Yaskawa INFORM job: LAB3-GROUPV2'2.JBI

/JOB
//NAME LAB3-GROUPV2'2
//POS
///NPOS 15,0,15,0,0,0
///TOOL 0
///POSTYPE PULSE
///PULSE
C00000=-729,-59979,-60060,-74,-89734,186
C00001=4452,18827,-51072,2986,-34195,44008
C00002=-2158,25887,-50796,2701,-28930,46142
C00003=-4327,35229,-34321,2660,-31477,21361
C00004=-13778,42742,-21333,8875,-39330,-13161
C00005=-15205,46983,-15261,9515,-46968,-18770
C00006=-16077,39808,-21056,7196,-36422,-13209
C00007=-21057,8484,-56828,1119,-11848,1649
C00008=-23284,14747,-79271,2827,22636,-7091
C00009=-18054,15511,-73334,806,11905,-7587
C00010=-19671,9683,-70517,8540,5629,-10803
C00011=-21717,17536,-102963,-1615,53770,-17043
C00012=-19881,21209,-97135,-2963,52531,-16955
C00013=-23771,9748,-100031,-181,45881,-17086
C00014=-1,-60103,-60032,2,-90053,2
EC00000=1
EC00001=-12851
EC00002=-12851
EC00003=-10530
EC00004=-2717
EC00005=-2717
EC00006=-22347
EC00007=-82435
EC00008=-82435
EC00009=-82435
EC00010=-82435
EC00011=-160520
EC00012=-160520
EC00013=-160520
EC00014=-1644
//INST
///DATE 2025/11/03 19:24
///ATTR SC,RW
///GROUP1 RB1,ST1
NOP
MOVJ C00000 EC00000 VJ=5.00
MOVJ C00001 EC00001 VJ=50.00
MOVC C00002 EC00002 V=83.3
ARCON ASF#(65)
MOVC C00003 EC00003
MOVC C00004 EC00004
MOVC C00005 EC00005 FPT
ARCOF AEF#(65)
MOVL C00006 EC00006 V=83.3
MOVJ C00007 EC00007 VJ=25.00
MOVL C00008 EC00008 V=83.3
ARCON ASF#(65)
MOVL C00009 EC00009
ARCOF AEF#(65)
MOVL C00010 EC00010 V=333.3
MOVL C00011 EC00011 V=50.0
ARCON ASF#(66)
MOVL C00012 EC00012
ARCOF AEF#(66)
MOVL C00013 EC00013 V=333.3
MOVJ C00014 EC00014 VJ=22.22
END
